Fanuc KAREL source: kb00193.KL

-- PROVISIONAL review KL for V1013-1; original PC SHA256 f361af43db382ea79e8cf2bc59fba775f00848deb2d4b58a2bcf06abc1a669b0
-- Incomplete behavior may be omitted. Consult companion uncertainty JSON. Do not deploy.
PROGRAM KB00193
%NOLOCKGROUP
BEGIN
  -- UNRESOLVED_PC offsets 5-12; opcodes 9D,23
  -- UNRESOLVED_PC offsets 17-24; opcodes 9D,23
  -- UNRESOLVED_PC offsets 29-45; opcodes 27,22,22,31
  -- UNRESOLVED_PC offsets 50-54; opcodes 7F
END KB00193
